Fanuc KAREL source: KO00054.KL

PROGRAM KO00054
%NOLOCKGROUP
%ENVIRONMENT MIR
VAR
  P1: XYZWPR
  P2: XYZWPR
  F: BOOLEAN
  OUT: XYZWPR
BEGIN
  F = TRUE
  OUT = MIRROR(P1, P2, F)
END KO00054
